Staubli VAL3: isReachable.pgx

public program isReachable(string x_sKey, num x_nIndex, tool x_tTool)
  local pointRx l_pPoint
  local bool l_bResult
  local mdesc l_mDesc
  local jointRx l_jJoint
begin
  if trajTemp:tTrajItem[x_sKey].pPointItem[x_nIndex].pParaItem.nMoveType==0
    l_mDesc=trajTemp:tTrajItem[x_sKey].pPointItem[x_nIndex].pParaItem.mMdesc
    l_pPoint.trsf=trajTemp:tTrajItem[x_sKey].pPointItem.pPointRx.trsf
    l_pPoint.config=trajTemp:tTrajItem[x_sKey].pPointItem.pPointRx.config
    l_bResult= pointToJoint(x_tTool,herej(),l_pPoint,l_jJoint)
    if l_bResult
      movel(l_pPoint,x_tTool,l_mDesc)
    endIf
  endIf
end
